# EPICS substitutions: db/Beckhoff_3XXX/ecmcEL3751.substitutions
file "ecmc_analogInputArray-chX.template"
{
  pattern {CH_ID, DTYP,                FTVL    }
          {01,    "asynInt32ArrayIn",  "LONG" }
}

file "ecmcEL3751_status-chX.template"
{
  pattern {CH_ID}
          {01   }
}

file "ecmc_controlWord-chX.template"
{
  pattern {CH_ID, KEY,   suffix,  sourceName, DESC             }
          {01,    "AI", "-Ctrl", "control",   "AI Control Word"}
}
